// TIA Portal V19 export
TYPE "PidL.Status"
   STRUCT
      OosAct : Bool;
      LocAct : Bool;
      ManAct : Bool;
      AutAct : Bool;
      SpExtAct : Bool;
      Protection : Bool;
      Intlock : Bool;
      Permit : Bool;
      TrackAct : Bool;
      SP : Real;
      PV : Real;
      ER : Real;
      MV : Real;
      PVOpScale : Struct
         High : Real;
         Low : Real;
      END_STRUCT;
      MVOpScale : Struct
         High : Real;
         Low : Real;
      END_STRUCT;
      SPIntLim : Struct
         High : Real;
         Low : Real;
      END_STRUCT;
      PV_unit : Int;
      MV_unit : Int;
   END_STRUCT;
END_TYPE
